Fanuc KAREL source: ka00012.KL

-- PROVISIONAL review KL for V1013-1; original PC SHA256 4ecfc04ca5ca17fe7501c48fc8340b1cc31edb8428c9d360c332152a202ff83f
-- Incomplete behavior may be omitted. Consult companion uncertainty JSON. Do not deploy.
PROGRAM KA00012
%NOLOCKGROUP
VAR
  SRC : INTEGER
-- UNRESOLVED_DECL DST type=002017
BEGIN
  -- UNRESOLVED_PC offsets 5-16; opcodes 2E,23
  -- UNRESOLVED_PC offsets 21-36; opcodes 21,22,9D,33,B4
  -- UNRESOLVED_PC offsets 41-45; opcodes 7F
END KA00012
